// TIA Portal V21 export
// export: Created 2026-11-10T19:12:21.8219882Z, ExportSetting WithDefaults, DisplayName Totally Integrated Automation Portal, DisplayVersion V21 Update 3, DisplayName STEP 7 Professional, DisplayVersion V21 Update 3, DisplayName STEP 7 Safety, DisplayVersion V21, DisplayName Tech WebApplication, DisplayVersion V21, DisplayName WinCC Basic/Comfort/Advanced, DisplayVersion V21 Update 3, DisplayName WinCC Unified, DisplayVersion V21 Update 3
DATA_BLOCK "DBsCONT_S"   // DB32
// stored: AutoNumber true, DBAccessibleFromOPCUA true, DBAccessibleFromWebserver true, InstanceOfName CONT_S, OfSystemLibElement CONT_S, OfSystemLibVersion 1.1
CONT_S   // technology object, version 1.1
   // VAR_INPUT
   //    COM_RST : Bool;
   //    LMNR_HS : Bool;
   //    LMNR_LS : Bool;
   //    LMNS_ON : Bool;
   //    LMNUP : Bool;
   //    LMNDN : Bool;
   //    PVPER_ON : Bool;
   //    CYCLE : Time;
   //    SP_INT : Real;
   //    PV_IN : Real;
   //    PV_PER : Word;
   //    GAIN : Real;
   //    TI : Time;
   //    DEADB_W : Real;
   //    PV_FAC : Real;
   //    PV_OFF : Real;
   //    PULSE_TM : Time;
   //    BREAK_TM : Time;
   //    MTR_TM : Time;
   //    DISV : Real;
   // END_VAR
   // VAR_OUTPUT
   //    QLMNUP : Bool;
   //    QLMNDN : Bool;
   //    PV : Real;
   //    ER : Real;
   // END_VAR
   // VAR RETAIN
   //    LMNRS_ON : Bool;
   //    LMNRSVAL : Real;
   //    LMNR_SIM : Real;
   //    sFbPVal : Real;
   //    sThrOn : Real;
   //    siImpAus : Int;
   //    stImpDauer : Time;
   //    stPausDauer : Time;
   // END_VAR
BEGIN
END_DATA_BLOCK
